FUNCTION_BLOCK FB_DosingPump EXTENDS FB_SFC_Cycle
VAR_INPUT
END_VAR
VAR_OUTPUT
	valve_A			: BOOL;
	valve_B			: BOOL;
END_VAR
VAR

	action_Time		: TIME:=T#0.5S;
	startDelay		: TIME:=T#0S;
	
	reqTiks			: DINT:=5;
	actTiks			: DINT:=5;
	
	fStageVolume	: REAL:=65; 	// CC/stage
	fReqVolume		: REAL:=500.0; 	// CC
	fActVolume		: REAL; 		// CC


END_VAR

VAR PERSISTENT
	
END_VAR

act_GetReference();

act_Oper();

reqTiks:=TRUNC(fReqVolume/fStageVolume);
fActVolume:=(actTiks*fStageVolume);

ACTION _acheck_Count_active:
bStepDone:=FALSE;
IF actTiks>=reqTiks THEN;
	bStepDone:=TRUE;
END_IF
END_ACTION

ACTION _acheck_Count_entry:
actTiks:=actTiks+1;
END_ACTION

ACTION _aDone_entry:
bRun:=FALSE;
bDone:=TRUE;
END_ACTION

ACTION _aInit_act_Oper_active:
SFCReset:=FALSE;
END_ACTION

ACTION _aInit_act_Oper_exit:
valve_A:=valve_B:=bRun:=bDone:=FALSE;
END_ACTION

ACTION _aReady_exit:
actTiks:=0;
END_ACTION

ACTION _astage_A_entry:
valve_A:=TRUE;
END_ACTION

ACTION _astage_A_exit:
valve_A:=FALSE;
END_ACTION

ACTION _astage_B_entry:
valve_B:=TRUE;
END_ACTION

ACTION _astage_B_exit:
valve_B:=FALSE;
END_ACTION

ACTION act_GetReference:
m_Set_SFCFlags_Reference();
END_ACTION

ACTION act_Oper:
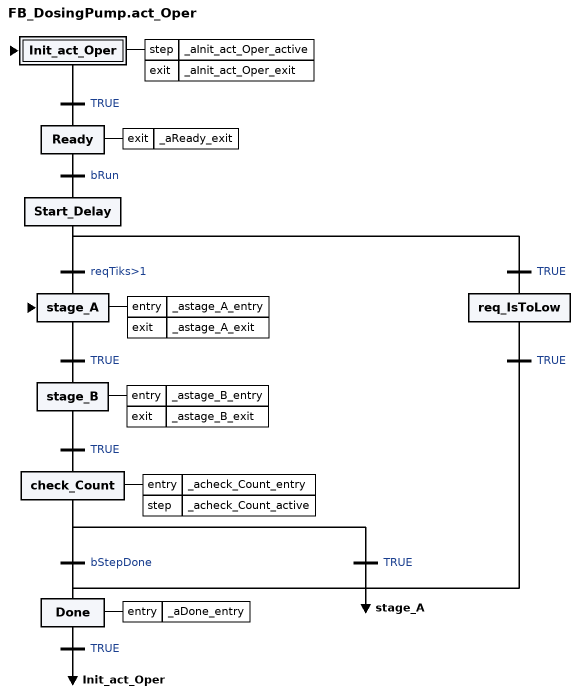
INITIAL_STEP Init_act_Oper:
    _aInit_act_Oper_active(N);  // step action
    _aInit_act_Oper_exit(P0);  // exit action
END_STEP
TRANSITION FROM Init_act_Oper TO Ready
    := TRUE;
END_TRANSITION
STEP Ready:
    _aReady_exit(P0);  // exit action
END_STEP
TRANSITION FROM Ready TO Start_Delay
    := bRun;
END_TRANSITION
STEP Start_Delay:  // min time startDelay
END_STEP
TRANSITION FROM Start_Delay TO stage_A
    := reqTiks>1;
END_TRANSITION
STEP stage_A:  // min time action_Time
    _astage_A_entry(P1);  // entry action
    _astage_A_exit(P0);  // exit action
END_STEP
TRANSITION FROM stage_A TO stage_B
    := TRUE;
END_TRANSITION
STEP stage_B:  // min time action_Time
    _astage_B_entry(P1);  // entry action
    _astage_B_exit(P0);  // exit action
END_STEP
TRANSITION FROM stage_B TO check_Count
    := TRUE;
END_TRANSITION
STEP check_Count:
    _acheck_Count_entry(P1);  // entry action
    _acheck_Count_active(N);  // step action
END_STEP
TRANSITION FROM check_Count TO Done
    := bStepDone;
END_TRANSITION
TRANSITION FROM check_Count TO stage_A
    := TRUE;
END_TRANSITION
TRANSITION FROM Start_Delay TO req_IsToLow
    := TRUE;
END_TRANSITION
STEP req_IsToLow:
END_STEP
TRANSITION FROM req_IsToLow TO Done
    := TRUE;
END_TRANSITION
STEP Done:
    _aDone_entry(P1);  // entry action
END_STEP
TRANSITION FROM Done TO Init_act_Oper
    := TRUE;
END_TRANSITION
// branch label Branch0_act_Oper
// branch label Branch1_act_Oper
END_ACTION

METHOD m_RunVolume : BOOL
VAR_INPUT
	Volume	:REAL;
END_VAR
fReqVolume:=Volume;
mRun();
IF rtDone.Q THEN;
	m_RunVolume:=TRUE;	
END_IF
END_METHOD

METHOD m_Set_SFCFlags_Reference : BOOL
//Set reference to SFC flags

refSFC.SFCInit REF= SFCInit;
refSFC.SFCReset REF= SFCReset;
refSFC.SFCError REF= SFCError;
refSFC.SFCEnableLimit REF= SFCEnableLimit;
refSFC.SFCErrorStep REF= SFCErrorStep;
refSFC.SFCErrorPOU REF= SFCErrorPOU;
refSFC.SFCQuitError REF= SFCQuitError;
refSFC.SFCPause REF= SFCPause;
refSFC.SFCTrans REF= SFCTrans;
refSFC.SFCCurrentStep REF= SFCCurrentStep;
refSFC.SFCTip REF= SFCTip;
refSFC.SFCTipMode REF= SFCTipMode;

// Cycle handle for SFC
m_SFC_Handle();
END_METHOD

METHOD m_Stop : BOOL
VAR_INPUT
END_VAR
SFCReset:=TRUE;
END_METHOD

END_FUNCTION_BLOCK

(* stored: Version 1.1.0.1, ProductVersion 3.1.4024.12
   POU FB_DosingPump: Id {7c08c2ba-d9cf-4bfb-abfd-8e2c5a78618b}, SpecialFunc None
   Folder manage: Id {f3c1175b-51b4-45b8-98a1-aa077b9febe6}
   Action _acheck_Count_active: Id {5ea15c14-afbb-4ed1-bc8c-231ae33b3975}
   Action _acheck_Count_entry: Id {3171b471-6b83-4f11-aa23-4f3b11832b2d}
   Action _aDone_entry: Id {5eab29f8-9325-48be-b604-8d8a46c98c66}
   Action _aInit_act_Oper_active: Id {dcd900aa-a12c-46e1-abde-573ca81c39da}
   Action _aInit_act_Oper_exit: Id {ee3e6fcb-aed9-4bc6-abb4-dfaefa95ae37}
   Action _aReady_exit: Id {6a2e8dc9-d34f-4af3-83cb-d604a06879bf}
   Action _astage_A_entry: Id {0f012b3f-8d5a-4f9c-9d7a-dc0e18fec8e8}
   Action _astage_A_exit: Id {c3b900d5-ebee-4d55-8b59-2af86500cbd9}
   Action _astage_B_entry: Id {aa4961fb-a8c3-4177-9ad3-c810d135bd77}
   Action _astage_B_exit: Id {b8b17864-ecbb-4f3e-a185-2a0cb2b44532}
   Action act_GetReference: Id {7d72703b-2334-4668-8865-0b9a7c7be4e3}
   Action act_Oper: Id {762d79ea-73b9-4b09-8d79-1296bfe123e6}
   Method m_RunVolume: Id {0d856e46-de18-4a27-9bfe-92513e0d3ab8}
   Method m_Set_SFCFlags_Reference: Id {b86dd4e2-3c28-4c4e-ac24-8fad9b06dbde}
   Method m_Stop: Id {a4b5a574-39b4-41ee-a2fd-a4f071a60b58} *)
